(* IEC 61131-3 sources: krc-sample-programs/motor-ramp-alarms-codesys/source/06_Programs, 4 files *)

(* ---- ALARMS.st ---- *)
PROGRAM ALARMS
VAR
	i            : INT;	// The alarm being looked at
	bAnyAlarm    : BOOL;	// Rollup while the list is scanned
	bAnyWarning  : BOOL;	// Rollup while the list is scanned
	bAnyUnacked  : BOOL;	// Rollup while the list is scanned
END_VAR
// ---- body ----
// ALARMS: times every step that waits on the machine, wires each alarm's trigger, and runs the alarm
// list. It runs after STATE_MACHINE, so it times the step the machine is in now. Reset is handled here: its
// press acknowledges the alarms, and once no ALARM-level alarm is left on the list, the state machine
// leaves Fault on its next scan.

// The step timeouts. If a step waits on the machine, it gets a timeout; if it waits on a person (Not
// Ready, Ready), it doesn't. Each timer runs only while its step is active, so it starts from zero
// every time the step starts.
TON_RAMP_10(IN := iStep = S4_RAMP_10, PT := T#1S * HMI_iRampTimeout);
TON_RAMP_25(IN := iStep = S4_RAMP_25, PT := T#1S * HMI_iRampTimeout);
TON_RAMP_50(IN := iStep = S4_RAMP_50, PT := T#1S * HMI_iRampTimeout);
TON_RAMP_75(IN := iStep = S4_RAMP_75, PT := T#1S * HMI_iRampTimeout);
TON_STOPPING(IN := iStep = S5_STOPPING, PT := T#1S * HMI_iStopTimeout);

// The speed feedback, watched the whole time the motor is at speed, not just on the way up: further off
// the reference than SPEED_DEVIATION, for T_SPEED_DEVIATION.
TON_SpeedDeviation(IN := iStep = S4_AT_SPEED AND ABS(iSpeedRef - iSpeedFbk) > SPEED_DEVIATION,
                   PT := T_SPEED_DEVIATION);

// Each alarm's trigger: one line each, the condition right now, written against the value it watches.
aAlarms[ALM_ESTOP].bTriggered := NOT bEStopOK;
aAlarms[ALM_DRIVE_DROPPED].bTriggered := NOT bDriveReady AND iStep >= S4_RAMP_10 AND iStep <= S5_STOPPING;
aAlarms[ALM_DRIVE_LOCAL].bTriggered := NOT bDriveRemote AND iStep >= S4_RAMP_10 AND iStep <= S5_STOPPING;
aAlarms[ALM_RAMP_TIMEOUT].bTriggered := (TON_RAMP_10.Q AND iSpeedFbk < SPEED_10)
                                     OR (TON_RAMP_25.Q AND iSpeedFbk < SPEED_25)
                                     OR (TON_RAMP_50.Q AND iSpeedFbk < SPEED_50)
                                     OR (TON_RAMP_75.Q AND iSpeedFbk < SPEED_75);
aAlarms[ALM_STOP_TIMEOUT].bTriggered := TON_STOPPING.Q AND iSpeedFbk > SPEED_STOPPED;
aAlarms[ALM_SPEED_DEVIATION].bTriggered := TON_SpeedDeviation.Q;
aAlarms[ALM_SIM_MODE].bTriggered := SIM_ENABLED;

// The alarm list. Every alarm lives the same way: it goes on the list when it triggers, the press of ACK
// or Reset acknowledges it, and it comes off once it is acknowledged AND its trigger is gone.
bAnyAlarm := FALSE;
bAnyWarning := FALSE;
bAnyUnacked := FALSE;
FOR i := 1 TO ALARM_COUNT DO
    // On: it triggered and isn't on the list yet. Not acknowledged, and it keeps the step it came on in
    // (the step the scan started in, before an override sent the machine to Fault).
    IF aAlarms[i].bTriggered AND NOT aAlarms[i].bOnList THEN
        aAlarms[i].bOnList := TRUE;
        aAlarms[i].bAcked := FALSE;
        aAlarms[i].iStepRaised := iStepAtScanStart;
    END_IF
    // Acknowledged: on the press of ACK or Reset (the one-shots).
    IF aAlarms[i].bOnList AND (rtAck.Q OR rtReset.Q) THEN
        aAlarms[i].bAcked := TRUE;
    END_IF
    // Off: acknowledged and the trigger gone.
    IF aAlarms[i].bOnList AND aAlarms[i].bAcked AND NOT aAlarms[i].bTriggered THEN
        aAlarms[i].bOnList := FALSE;
    END_IF
    // What the rest of the program needs to know about the list.
    bAnyAlarm := bAnyAlarm OR (aAlarms[i].bOnList AND aAlarms[i].eLevel = LVL_ALARM);
    bAnyWarning := bAnyWarning OR (aAlarms[i].bOnList AND aAlarms[i].eLevel = LVL_WARNING);
    bAnyUnacked := bAnyUnacked OR (aAlarms[i].bOnList AND NOT aAlarms[i].bAcked AND aAlarms[i].eLevel >= LVL_WARNING);
END_FOR
bAlarmOnList := bAnyAlarm;
bWarningOnList := bAnyWarning;
bUnacknowledged := bAnyUnacked;

(* ---- DEVICES.st ---- *)
PROGRAM DEVICES
// ---- body ----
// DEVICES: every output is set here, once, from the step, like a coil: assigned its condition every scan,
// TRUE while the condition is true and FALSE as soon as it isn't.

// The permissives: one line each, what each one waits for.
aPermissives[PERM_DRIVE_READY].bSatisfied := bDriveReady;
aPermissives[PERM_DRIVE_REMOTE].bSatisfied := bDriveRemote;
aPermissives[PERM_STOP_RELEASED].bSatisfied := NOT bStopPB;
aPermissives[PERM_MOTOR_STOPPED].bSatisfied := iSpeedFbk <= SPEED_STOPPED;

// Motor run: on while running and while stopping, so the drive brings the motor down under control.
bMotorRun := iStep >= S4_RAMP_10 AND iStep <= S5_STOPPING;

// Speed reference: one CASE, so it is written in one place and every step gets a value.
CASE iStep OF
S4_RAMP_10:
    iSpeedRef := SPEED_10;
S4_RAMP_25:
    iSpeedRef := SPEED_25;
S4_RAMP_50:
    iSpeedRef := SPEED_50;
S4_RAMP_75, S4_AT_SPEED:
    iSpeedRef := SPEED_75;
ELSE
    iSpeedRef := 0;
END_CASE

// Stack light green: running.
bStackGreen := iStep >= S4_RAMP_10 AND iStep <= S4_AT_SPEED;

// Stack light red: not running. Written from the steps, never from another output.
bStackRed := iStep < S4_RAMP_10 OR iStep >= S5_STOPPING;

// The flasher: a timer that restarts itself. Its done bit is on for one scan every T_FLASH, and each
// time it is, the flash flips.
TON_Flash(IN := NOT TON_Flash.Q, PT := T_FLASH);
IF TON_Flash.Q THEN
    bFlash := NOT bFlash;
END_IF

// Stack light orange, the alarm light: flashing while an alarm or warning hasn't been acknowledged,
// steady while one is still on the list.
bStackOrange := (bUnacknowledged AND bFlash) OR ((bAlarmOnList OR bWarningOnList) AND NOT bUnacknowledged);

// The button lamps: lit when the button can be pressed.
bStartLamp := iStep = S3_READY;
bStopLamp := iStep >= S4_RAMP_10 AND iStep <= S4_AT_SPEED;
bResetLamp := iStep = S6_FAULT;
bAckLamp := bUnacknowledged;

(* ---- OUTPUTS.st ---- *)
PROGRAM OUTPUTS
VAR
	i       : INT;	// The line, or the alarm, being looked at
	iLines  : INT;	// How many alarms are on the list, up to ALARM_LINES
	aShown  : ARRAY[1..ALARM_LINES] OF INT;	// Which alarm each line shows
	sLevel  : STRING(10);	// The line's level, in words
END_VAR
// ---- body ----
// OUTPUTS: every output is written here and nowhere else. First the hardware, in terminal order.
DO_bMotorRun := bMotorRun;
DO_bStackGreen := bStackGreen;
DO_bStackRed := bStackRed;
DO_bStackOrange := bStackOrange;

// Speed reference to the drive: 0 to 100 % becomes 0 to 32767 (AO_FULL_SCALE), 0 to 10 V, rounded to the
// nearest count.
AO_wSpeedRef := DINT_TO_WORD((INT_TO_DINT(iSpeedRef) * AO_FULL_SCALE + 50) / 100);

// Then the HMI. The screen only reads these.
HMI_bStartLamp := bStartLamp;
HMI_bStopLamp := bStopLamp;
HMI_bResetLamp := bResetLamp;
HMI_bAckLamp := bAckLamp;
HMI_bStackGreen := bStackGreen;
HMI_bStackOrange := bStackOrange;
HMI_bStackRed := bStackRed;
HMI_bMotorRun := bMotorRun;
HMI_iSpeedRef := iSpeedRef;
HMI_iSpeedFbk := iSpeedFbk;
HMI_sState := sStateDescription;

// The permissive lamps.
FOR i := 1 TO PERMISSIVE_COUNT DO
    HMI_abPermissive[i] := aPermissives[i].bSatisfied;
END_FOR

// The alarm lines: the alarms on the list, in table order (ALARM level first), up to ALARM_LINES. Each
// line is the level, the words, and the step the machine was in when it came on.
iLines := 0;
FOR i := 1 TO ALARM_COUNT DO
    IF aAlarms[i].bOnList AND iLines < ALARM_LINES THEN
        iLines := iLines + 1;
        aShown[iLines] := i;
    END_IF
END_FOR
FOR i := 1 TO ALARM_LINES DO
    IF i <= iLines THEN
        CASE aAlarms[aShown[i]].eLevel OF
        LVL_ALARM:
            sLevel := 'ALARM';
        LVL_WARNING:
            sLevel := 'WARNING';
        ELSE
            sLevel := 'INFO';
        END_CASE
        HMI_asAlarmLine[i] := CONCAT(CONCAT(sLevel, '   '), CONCAT(aAlarms[aShown[i]].sText,
                              CONCAT('   (step ', CONCAT(INT_TO_STRING(aAlarms[aShown[i]].iStepRaised), ')'))));
        HMI_abAlarmUnacked[i] := NOT aAlarms[aShown[i]].bAcked;
    ELSE
        HMI_asAlarmLine[i] := '';
        HMI_abAlarmUnacked[i] := FALSE;
    END_IF
END_FOR

(* ---- STATE_MACHINE.st ---- *)
PROGRAM STATE_MACHINE
VAR
	i            : INT;	// The permissive being looked at
	bAllMet      : BOOL;	// Rollup while the permissives are scanned
	sWaitingFor  : STRING(30);	// The first permissive not met
END_VAR
// ---- body ----
// STATE_MACHINE: decides which step the machine is in. The steps are the values of the enum E_Step
// (03_States). iStep is the step the machine is in; each exit puts the next step into iNextStep, and the
// step only changes on the last line, so every line in one scan sees the same step.

// The permissives: everything Ready waits for, one line each in the permissive table (GVL_Alarms), each
// wired in DEVICES. This rollup ANDs them, and keeps the first one not met so Not Ready can name it.
bAllMet := TRUE;
sWaitingFor := '';
FOR i := 1 TO PERMISSIVE_COUNT DO
    IF bAllMet AND NOT aPermissives[i].bSatisfied THEN
        sWaitingFor := aPermissives[i].sText;
    END_IF
    bAllMet := bAllMet AND aPermissives[i].bSatisfied;
END_FOR
bPermissivesOK := bAllMet;

// Every state writes what it is doing, in words, for the screen.
CASE iStep OF

S0_IDLE:
    // Idle: powered up and at rest. Go to Not Ready.
    sStateDescription := 'Idle';
    iNextStep := S1_NOT_READY;

S1_NOT_READY:
    // Not Ready never just says Not Ready: it names the first permissive it is waiting for.
    IF bPermissivesOK THEN
        sStateDescription := 'Not Ready - every permissive met';
    ELSE
        sStateDescription := CONCAT('Not Ready - waiting for: ', sWaitingFor);
    END_IF
    // Every permissive met: ready.
    IF bPermissivesOK THEN
        iNextStep := S3_READY;
    END_IF

S3_READY:
    sStateDescription := 'Ready - press Start';
    // Start pressed: the one-shot, so a held Start doesn't count. Start the motor at 10 %.
    IF rtStart.Q THEN
        iNextStep := S4_RAMP_10;
    END_IF
    // A permissive dropped: back to Not Ready, which says which one. Last, so it wins over Start.
    IF NOT bPermissivesOK THEN
        iNextStep := S1_NOT_READY;
    END_IF

S4_RAMP_10:
    sStateDescription := 'Running - ramping to 10 %';
    // The speed feedback has reached 10 %: next step. Its timeout is an alarm now (ALARMS).
    IF iSpeedFbk >= SPEED_10 THEN
        iNextStep := S4_RAMP_25;
    END_IF

S4_RAMP_25:
    sStateDescription := 'Running - ramping to 25 %';
    IF iSpeedFbk >= SPEED_25 THEN
        iNextStep := S4_RAMP_50;
    END_IF

S4_RAMP_50:
    sStateDescription := 'Running - ramping to 50 %';
    IF iSpeedFbk >= SPEED_50 THEN
        iNextStep := S4_RAMP_75;
    END_IF

S4_RAMP_75:
    sStateDescription := 'Running - ramping to 75 %';
    IF iSpeedFbk >= SPEED_75 THEN
        iNextStep := S4_AT_SPEED;
    END_IF

S4_AT_SPEED:
    // At speed: no exit of its own. It holds here until Stop, below.
    sStateDescription := 'Running - at speed, 75 %';

S5_STOPPING:
    sStateDescription := 'Stopping - waiting for the motor to stop';
    // The motor has stopped. Back to Not Ready.
    IF iSpeedFbk <= SPEED_STOPPED THEN
        iNextStep := S1_NOT_READY;
    END_IF

S6_FAULT:
    // Fault: the alarm list says why. The state machine carries no alarm text, only what it is doing.
    sStateDescription := 'Fault - see the alarm list, then press Reset';
    // Reset is handled in ALARMS: its press tries to clear every latched alarm. One whose cause is gone
    // comes off the list; one still latched means its fault is still active. Once no ALARM-level alarm is
    // left, Fault is over: straight to Not Ready, which checks every permissive again before Ready.
    IF NOT bAlarmOnList THEN
        iNextStep := S1_NOT_READY;
    END_IF

ELSE
    // A step that isn't in the list can't happen, but if it ever does, fail safe.
    sStateDescription := 'Fault - unknown step';
    iNextStep := S6_FAULT;
END_CASE

// Stop, out of any running step: written once for the whole Running state, not in every ramp step.
IF iStep >= S4_RAMP_10 AND iStep <= S4_AT_SPEED AND bStopPB THEN
    iNextStep := S5_STOPPING;
END_IF

// The global overrides, after everything else, so they always win the scan.
// 1. The E-stop circuit is open.
IF NOT bEStopOK THEN
    iNextStep := S6_FAULT;
END_IF
// 2. An ALARM-level alarm is on the list. It holds the machine in Fault until it is acknowledged and gone.
IF bAlarmOnList THEN
    iNextStep := S6_FAULT;
END_IF

// Take the next step. This is the only place the step changes. ALARMS runs after this, so keep the step
// the scan started in: an alarm's line names where the machine was, not the Fault it was just sent to.
iStepAtScanStart := iStep;
iStep := iNextStep;
